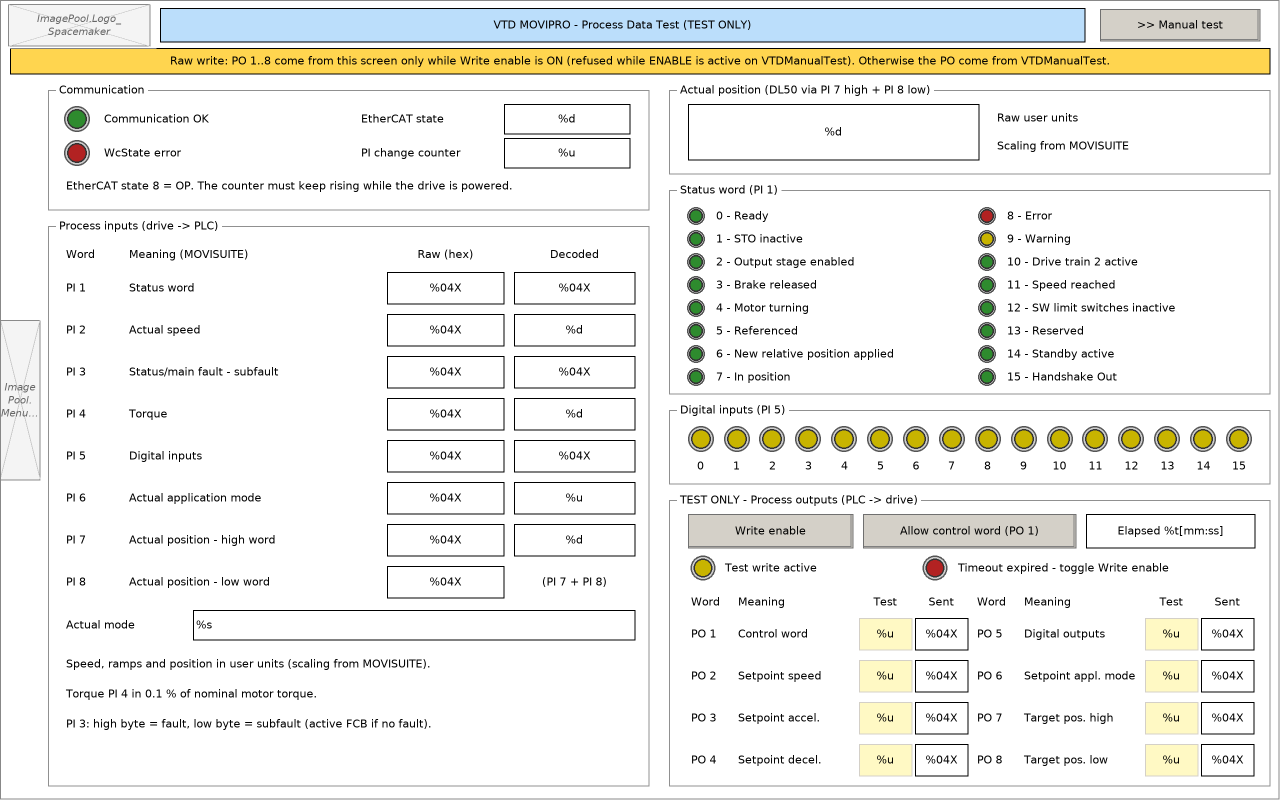
VISUALIZATION Visualization  // 1280x800
    GroupBox (48,82 601x128), "Communication"
    GroupBox (48,218 601x568), "Process inputs (drive -> PLC)"
    GroupBox (669,82 601x92), "Actual position (DL50 via PI 7 high + PI 8 low)"
    GroupBox (669,182 601x212), "Status word (PI 1)"
    GroupBox (669,402 601x82), "Digital inputs (PI 5)"
    GroupBox (669,492 601x294), "TEST ONLY - Process outputs (PLC -> drive)"
    Rectangle (160,8 925x34), "VTD MOVIPRO - Process Data Test (TEST ONLY)"
    Rectangle (10,48 1260x26), "Raw write: PO 1..8 come from this screen only while Write enable is ON (refused while ENABLE is active on VTDManualTest). Otherwise the PO come from VTDManualTest."
    Lamp1 (62,104 30x30), variable: GVL_HMI_VTD.stPdStatus.bCommunicationOk, style: Lamp-Lamp1-Green
    Rectangle (101,104 243x30), "Communication OK"
    Lamp1 (62,138 30x30), variable: GVL_HMI_VTD.stPdStatus.bWcStateError, style: Lamp-Lamp1-Red
    Rectangle (101,138 243x30), "WcState error"
    Rectangle (358,104 146x30), "EtherCAT state"
    Rectangle (504,104 126x30), "%d", text variable: GVL_HMI_VTD.stPdStatus.uiEcState
    Rectangle (358,138 146x30), "PI change counter"
    Rectangle (504,138 126x30), "%u", text variable: GVL_HMI_VTD.stPdStatus.udiInputChangeCount
    Rectangle (63,172 572x28), "EtherCAT state 8 = OP. The counter must keep rising while the drive is powered."
    Rectangle (63,242 58x25), "Word"
    Rectangle (126,242 252x25), "Meaning (MOVISUITE)"
    Rectangle (387,242 117x25), "Raw (hex)"
    Rectangle (514,242 121x25), "Decoded"
    Rectangle (63,272 58x32), "PI 1"
    Rectangle (126,272 252x32), "Status word"
    Rectangle (387,272 117x32), "%04X", text variable: GVL_HMI_VTD.stPdStatus.aProcessInputRaw[1]
    Rectangle (514,272 121x32), "%04X", text variable: GVL_HMI_VTD.stPdStatus.wStatusWord
    Rectangle (63,314 58x32), "PI 2"
    Rectangle (126,314 252x32), "Actual speed"
    Rectangle (387,314 117x32), "%04X", text variable: GVL_HMI_VTD.stPdStatus.aProcessInputRaw[2]
    Rectangle (514,314 121x32), "%d", text variable: GVL_HMI_VTD.stPdStatus.iActualSpeedRaw
    Rectangle (63,356 58x32), "PI 3"
    Rectangle (126,356 252x32), "Status/main fault - subfault"
    Rectangle (387,356 117x32), "%04X", text variable: GVL_HMI_VTD.stPdStatus.aProcessInputRaw[3]
    Rectangle (514,356 121x32), "%04X", text variable: GVL_HMI_VTD.stPdStatus.wFaultCode
    Rectangle (63,398 58x32), "PI 4"
    Rectangle (126,398 252x32), "Torque"
    Rectangle (387,398 117x32), "%04X", text variable: GVL_HMI_VTD.stPdStatus.aProcessInputRaw[4]
    Rectangle (514,398 121x32), "%d", text variable: GVL_HMI_VTD.stPdStatus.iTorqueRaw
    Rectangle (63,440 58x32), "PI 5"
    Rectangle (126,440 252x32), "Digital inputs"
    Rectangle (387,440 117x32), "%04X", text variable: GVL_HMI_VTD.stPdStatus.aProcessInputRaw[5]
    Rectangle (514,440 121x32), "%04X", text variable: GVL_HMI_VTD.stPdStatus.wDigitalInputs
    Rectangle (63,482 58x32), "PI 6"
    Rectangle (126,482 252x32), "Actual application mode"
    Rectangle (387,482 117x32), "%04X", text variable: GVL_HMI_VTD.stPdStatus.aProcessInputRaw[6]
    Rectangle (514,482 121x32), "%u", text variable: GVL_HMI_VTD.stPdStatus.uiActualApplicationMode
    Rectangle (63,524 58x32), "PI 7"
    Rectangle (126,524 252x32), "Actual position - high word"
    Rectangle (387,524 117x32), "%04X", text variable: GVL_HMI_VTD.stPdStatus.aProcessInputRaw[7]
    Rectangle (514,524 121x32), "%d", text variable: GVL_HMI_VTD.stPdStatus.diActualPositionRaw
    Rectangle (63,566 58x32), "PI 8"
    Rectangle (126,566 252x32), "Actual position - low word"
    Rectangle (387,566 117x32), "%04X", text variable: GVL_HMI_VTD.stPdStatus.aProcessInputRaw[8]
    Rectangle (514,566 121x32), "(PI 7 + PI 8)"
    Rectangle (63,610 126x30), "Actual mode"
    Rectangle (193,610 442x30), "%s", text variable: GVL_HMI_VTD.stPdStatus.sActualModeName
    Rectangle (63,650 572x28), "Speed, ramps and position in user units (scaling from MOVISUITE)."
    Rectangle (63,680 572x28), "Torque PI 4 in 0.1 % of nominal motor torque."
    Rectangle (63,710 572x28), "PI 3: high byte = fault, low byte = subfault (active FCB if no fault)."
    Rectangle (688,104 291x56), "%d", text variable: GVL_HMI_VTD.stPdStatus.diActualPositionRaw
    Rectangle (994,104 261x28), "Raw user units"
    Rectangle (994,132 261x28), "Scaling from MOVISUITE"
    Lamp1 (686,206 20x20), variable: GVL_HMI_VTD.stPdStatus.wStatusWord.0, style: Lamp-Lamp1-Green
    Rectangle (713,205 262x22), "0 - Ready"
    Lamp1 (686,229 20x20), variable: GVL_HMI_VTD.stPdStatus.wStatusWord.1, style: Lamp-Lamp1-Green
    Rectangle (713,228 262x22), "1 - STO inactive"
    Lamp1 (686,252 20x20), variable: GVL_HMI_VTD.stPdStatus.wStatusWord.2, style: Lamp-Lamp1-Green
    Rectangle (713,251 262x22), "2 - Output stage enabled"
    Lamp1 (686,275 20x20), variable: GVL_HMI_VTD.stPdStatus.wStatusWord.3, style: Lamp-Lamp1-Green
    Rectangle (713,274 262x22), "3 - Brake released"
    Lamp1 (686,298 20x20), variable: GVL_HMI_VTD.stPdStatus.wStatusWord.4, style: Lamp-Lamp1-Green
    Rectangle (713,297 262x22), "4 - Motor turning"
    Lamp1 (686,321 20x20), variable: GVL_HMI_VTD.stPdStatus.wStatusWord.5, style: Lamp-Lamp1-Green
    Rectangle (713,320 262x22), "5 - Referenced"
    Lamp1 (686,344 20x20), variable: GVL_HMI_VTD.stPdStatus.wStatusWord.6, style: Lamp-Lamp1-Green
    Rectangle (713,343 262x22), "6 - New relative position applied"
    Lamp1 (686,367 20x20), variable: GVL_HMI_VTD.stPdStatus.wStatusWord.7, style: Lamp-Lamp1-Green
    Rectangle (713,366 262x22), "7 - In position"
    Lamp1 (977,206 20x20), variable: GVL_HMI_VTD.stPdStatus.wStatusWord.8, style: Lamp-Lamp1-Red
    Rectangle (1004,205 262x22), "8 - Error"
    Lamp1 (977,229 20x20), variable: GVL_HMI_VTD.stPdStatus.wStatusWord.9, style: Lamp-Lamp1-Yellow
    Rectangle (1004,228 262x22), "9 - Warning"
    Lamp1 (977,252 20x20), variable: GVL_HMI_VTD.stPdStatus.wStatusWord.10, style: Lamp-Lamp1-Green
    Rectangle (1004,251 262x22), "10 - Drive train 2 active"
    Lamp1 (977,275 20x20), variable: GVL_HMI_VTD.stPdStatus.wStatusWord.11, style: Lamp-Lamp1-Green
    Rectangle (1004,274 262x22), "11 - Speed reached"
    Lamp1 (977,298 20x20), variable: GVL_HMI_VTD.stPdStatus.wStatusWord.12, style: Lamp-Lamp1-Green
    Rectangle (1004,297 262x22), "12 - SW limit switches inactive"
    Lamp1 (977,321 20x20), variable: GVL_HMI_VTD.stPdStatus.wStatusWord.13, style: Lamp-Lamp1-Green
    Rectangle (1004,320 262x22), "13 - Reserved"
    Lamp1 (977,344 20x20), variable: GVL_HMI_VTD.stPdStatus.wStatusWord.14, style: Lamp-Lamp1-Green
    Rectangle (1004,343 262x22), "14 - Standby active"
    Lamp1 (977,367 20x20), variable: GVL_HMI_VTD.stPdStatus.wStatusWord.15, style: Lamp-Lamp1-Green
    Rectangle (1004,366 262x22), "15 - Handshake Out"
    Lamp1 (686,424 30x30), variable: GVL_HMI_VTD.stPdStatus.wDigitalInputs.0, style: Lamp-Lamp1-Yellow
    Rectangle (686,456 29x20), "0"
    Lamp1 (722,424 30x30), variable: GVL_HMI_VTD.stPdStatus.wDigitalInputs.1, style: Lamp-Lamp1-Yellow
    Rectangle (722,456 29x20), "1"
    Lamp1 (757,424 30x30), variable: GVL_HMI_VTD.stPdStatus.wDigitalInputs.2, style: Lamp-Lamp1-Yellow
    Rectangle (758,456 29x20), "2"
    Lamp1 (793,424 30x30), variable: GVL_HMI_VTD.stPdStatus.wDigitalInputs.3, style: Lamp-Lamp1-Yellow
    Rectangle (794,456 29x20), "3"
    Lamp1 (829,424 30x30), variable: GVL_HMI_VTD.stPdStatus.wDigitalInputs.4, style: Lamp-Lamp1-Yellow
    Rectangle (830,456 29x20), "4"
    Lamp1 (865,424 30x30), variable: GVL_HMI_VTD.stPdStatus.wDigitalInputs.5, style: Lamp-Lamp1-Yellow
    Rectangle (866,456 29x20), "5"
    Lamp1 (901,424 30x30), variable: GVL_HMI_VTD.stPdStatus.wDigitalInputs.6, style: Lamp-Lamp1-Yellow
    Rectangle (901,456 30x20), "6"
    Lamp1 (937,424 30x30), variable: GVL_HMI_VTD.stPdStatus.wDigitalInputs.7, style: Lamp-Lamp1-Yellow
    Rectangle (937,456 29x20), "7"
    Lamp1 (973,424 30x30), variable: GVL_HMI_VTD.stPdStatus.wDigitalInputs.8, style: Lamp-Lamp1-Yellow
    Rectangle (973,456 29x20), "8"
    Lamp1 (1009,424 30x30), variable: GVL_HMI_VTD.stPdStatus.wDigitalInputs.9, style: Lamp-Lamp1-Yellow
    Rectangle (1009,456 29x20), "9"
    Lamp1 (1045,424 30x30), variable: GVL_HMI_VTD.stPdStatus.wDigitalInputs.10, style: Lamp-Lamp1-Yellow
    Rectangle (1045,456 29x20), "10"
    Lamp1 (1080,424 30x30), variable: GVL_HMI_VTD.stPdStatus.wDigitalInputs.11, style: Lamp-Lamp1-Yellow
    Rectangle (1081,456 29x20), "11"
    Lamp1 (1116,424 30x30), variable: GVL_HMI_VTD.stPdStatus.wDigitalInputs.12, style: Lamp-Lamp1-Yellow
    Rectangle (1117,456 29x20), "12"
    Lamp1 (1152,424 30x30), variable: GVL_HMI_VTD.stPdStatus.wDigitalInputs.13, style: Lamp-Lamp1-Yellow
    Rectangle (1153,456 29x20), "13"
    Lamp1 (1188,424 30x30), variable: GVL_HMI_VTD.stPdStatus.wDigitalInputs.14, style: Lamp-Lamp1-Yellow
    Rectangle (1189,456 29x20), "14"
    Lamp1 (1224,424 30x30), variable: GVL_HMI_VTD.stPdStatus.wDigitalInputs.15, style: Lamp-Lamp1-Yellow
    Rectangle (1224,456 30x20), "15"
    Button (688,514 165x34), "Write enable", colour toggle: GVL_HMI_VTD.stPdCommand.bTestWriteEnable
        toggle GVL_HMI_VTD.stPdCommand.bTestWriteEnable
    Button (863,514 213x34), "Allow control word (PO 1)", colour toggle: GVL_HMI_VTD.stPdCommand.bTestAllowControlWord, input disabled if: NOT GVL_HMI_VTD.stPdCommand.bTestWriteEnable
        toggle GVL_HMI_VTD.stPdCommand.bTestAllowControlWord
    Rectangle (1086,514 169x34), "Elapsed %t[mm:ss]", text variable: GVL_HMI_VTD.stPdStatus.tTestWriteElapsed
    Lamp1 (688,554 30x28), variable: GVL_HMI_VTD.stPdStatus.bTestWriteActive, style: Lamp-Lamp1-Yellow
    Rectangle (722,554 194x28), "Test write active"
    Lamp1 (920,554 30x28), variable: GVL_HMI_VTD.stPdStatus.bTestWriteExpired, style: Lamp-Lamp1-Red
    Rectangle (955,554 300x28), "Timeout expired - toggle Write enable"
    Rectangle (688,590 44x24), "Word"
    Rectangle (735,590 121x24), "Meaning"
    Rectangle (859,590 53x24), "Test"
    Rectangle (915,590 53x24), "Sent"
    Rectangle (688,618 44x32), "PO 1"
    Rectangle (735,618 121x32), "Control word"
    Textfield (859,618 53x32), "%u", text variable: GVL_HMI_VTD.stPdCommand.aTestProcessOutput[1], input disabled if: NOT GVL_HMI_VTD.stPdCommand.bTestAllowControlWord
        OnMouseClick: write the text variable via VisuDialogs.Numpad, min 0, max 65535
    Rectangle (915,618 53x32), "%04X", text variable: GVL_HMI_VTD.stPdStatus.aProcessOutputSent[1]
    Rectangle (688,660 44x32), "PO 2"
    Rectangle (735,660 121x32), "Setpoint speed"
    Textfield (859,660 53x32), "%u", text variable: GVL_HMI_VTD.stPdCommand.aTestProcessOutput[2]
        OnMouseClick: write the text variable via VisuDialogs.Numpad, min 0, max 65535
    Rectangle (915,660 53x32), "%04X", text variable: GVL_HMI_VTD.stPdStatus.aProcessOutputSent[2]
    Rectangle (688,702 44x32), "PO 3"
    Rectangle (735,702 121x32), "Setpoint accel."
    Textfield (859,702 53x32), "%u", text variable: GVL_HMI_VTD.stPdCommand.aTestProcessOutput[3]
        OnMouseClick: write the text variable via VisuDialogs.Numpad, min 0, max 65535
    Rectangle (915,702 53x32), "%04X", text variable: GVL_HMI_VTD.stPdStatus.aProcessOutputSent[3]
    Rectangle (688,744 44x32), "PO 4"
    Rectangle (735,744 121x32), "Setpoint decel."
    Textfield (859,744 53x32), "%u", text variable: GVL_HMI_VTD.stPdCommand.aTestProcessOutput[4]
        OnMouseClick: write the text variable via VisuDialogs.Numpad, min 0, max 65535
    Rectangle (915,744 53x32), "%04X", text variable: GVL_HMI_VTD.stPdStatus.aProcessOutputSent[4]
    Rectangle (974,590 44x24), "Word"
    Rectangle (1021,590 121x24), "Meaning"
    Rectangle (1145,590 53x24), "Test"
    Rectangle (1201,590 53x24), "Sent"
    Rectangle (974,618 44x32), "PO 5"
    Rectangle (1021,618 121x32), "Digital outputs"
    Textfield (1145,618 53x32), "%u", text variable: GVL_HMI_VTD.stPdCommand.aTestProcessOutput[5]
        OnMouseClick: write the text variable via VisuDialogs.Numpad, min 0, max 65535
    Rectangle (1201,618 53x32), "%04X", text variable: GVL_HMI_VTD.stPdStatus.aProcessOutputSent[5]
    Rectangle (974,660 44x32), "PO 6"
    Rectangle (1021,660 121x32), "Setpoint appl. mode"
    Textfield (1145,660 53x32), "%u", text variable: GVL_HMI_VTD.stPdCommand.aTestProcessOutput[6]
        OnMouseClick: write the text variable via VisuDialogs.Numpad, min 0, max 65535
    Rectangle (1201,660 53x32), "%04X", text variable: GVL_HMI_VTD.stPdStatus.aProcessOutputSent[6]
    Rectangle (974,702 44x32), "PO 7"
    Rectangle (1021,702 121x32), "Target pos. high"
    Textfield (1145,702 53x32), "%u", text variable: GVL_HMI_VTD.stPdCommand.aTestProcessOutput[7]
        OnMouseClick: write the text variable via VisuDialogs.Numpad, min 0, max 65535
    Rectangle (1201,702 53x32), "%04X", text variable: GVL_HMI_VTD.stPdStatus.aProcessOutputSent[7]
    Rectangle (974,744 44x32), "PO 8"
    Rectangle (1021,744 121x32), "Target pos. low"
    Textfield (1145,744 53x32), "%u", text variable: GVL_HMI_VTD.stPdCommand.aTestProcessOutput[8]
        OnMouseClick: write the text variable via VisuDialogs.Numpad, min 0, max 65535
    Rectangle (1201,744 53x32), "%04X", text variable: GVL_HMI_VTD.stPdStatus.aProcessOutputSent[8]
    Button (1100,9 160x32), ">> Manual test"
        OnMouseClick: change screen: VTDManualTest
    Rectangle (0,0 156x48)
        OnMouseClick: change screen: Main
    Image (8,4 142x42), image: ImagePool.Logo_Spacemaker
        OnMouseClick: change screen: Main
    Rectangle (0,320 40x160)
        OnMouseEnter: OpenDialog Dialog=Dialog, OpenModal=True, PositionX=0, PositionY=0
        OnMouseClick: OpenDialog Dialog=Dialog, OpenModal=True, PositionX=0, PositionY=0
    Image (0,320 40x160), image: ImagePool.Menu_Tab
        OnMouseEnter: OpenDialog Dialog=Dialog, OpenModal=True, PositionX=0, PositionY=0
        OnMouseClick: OpenDialog Dialog=Dialog, OpenModal=True, PositionX=0, PositionY=0
END_VISUALIZATION

(* stored: Version 1.1.0.1
   Visu Visualization: Id {042c51d0-c84f-427f-9fe7-9915de0e56a0} *)
